Fanuc KAREL source: KT00869.KL

PROGRAM KT00869
%NOLOCKGROUP
VAR
  I1: INTEGER
  I2: INTEGER
  OUT: REAL
BEGIN
  I1 = 2
  I2 = 3
  I1 = 2
  I2 = 3
  OUT = TRUNC(I1)
END KT00869
